Fanuc KAREL source: ke00002.KL

-- PROVISIONAL review KL for V1013-1; original PC SHA256 d42c953c20f10ee6536fb5e6948249b2925b12db68e7b335321004d960312c13
-- Incomplete behavior may be omitted. Consult companion uncertainty JSON. Do not deploy.
PROGRAM KE00002
%NOLOCKGROUP
BEGIN
  -- UNRESOLVED_PC offsets 5-17; opcodes 3F,75
  -- UNRESOLVED_PC offsets 22-29; opcodes 9D,23
  -- UNRESOLVED_PC offsets 34-46; opcodes 3F,22,9D,33,61
  -- UNRESOLVED_PC offsets 51-87; opcodes 27,22,2A,22,22,22,22,31
  -- UNRESOLVED_PC offsets 92-96; opcodes 7F
END KE00002
